// CFC twin of T_SafeTof_Tests: the same tests drawn as CFC diagrams, the way a TwinSAFE project is authored.
    FUNCTION_BLOCK T_SafeTof_Tests_CFC EXTENDS T_SafeCfcTestSuite
    VAR
    // Test_OutputDelayedOff
    group_1 : T_SafeGroup;
    fb_1 : T_SafeTof(group := group_1) := (Parameters := (DelayTime := T#100MS));
    trigStart_1 : R_TRIG;
    t0_1 : TON;
    t1_1 : TON;
    trig0_1 : R_TRIG;
    trig1_1 : R_TRIG;
END_VAR

Test_OutputDelayedOff();

METHOD PRIVATE Test_OutputDelayedOff
// note: this text did not pass the execution check against the stored diagram
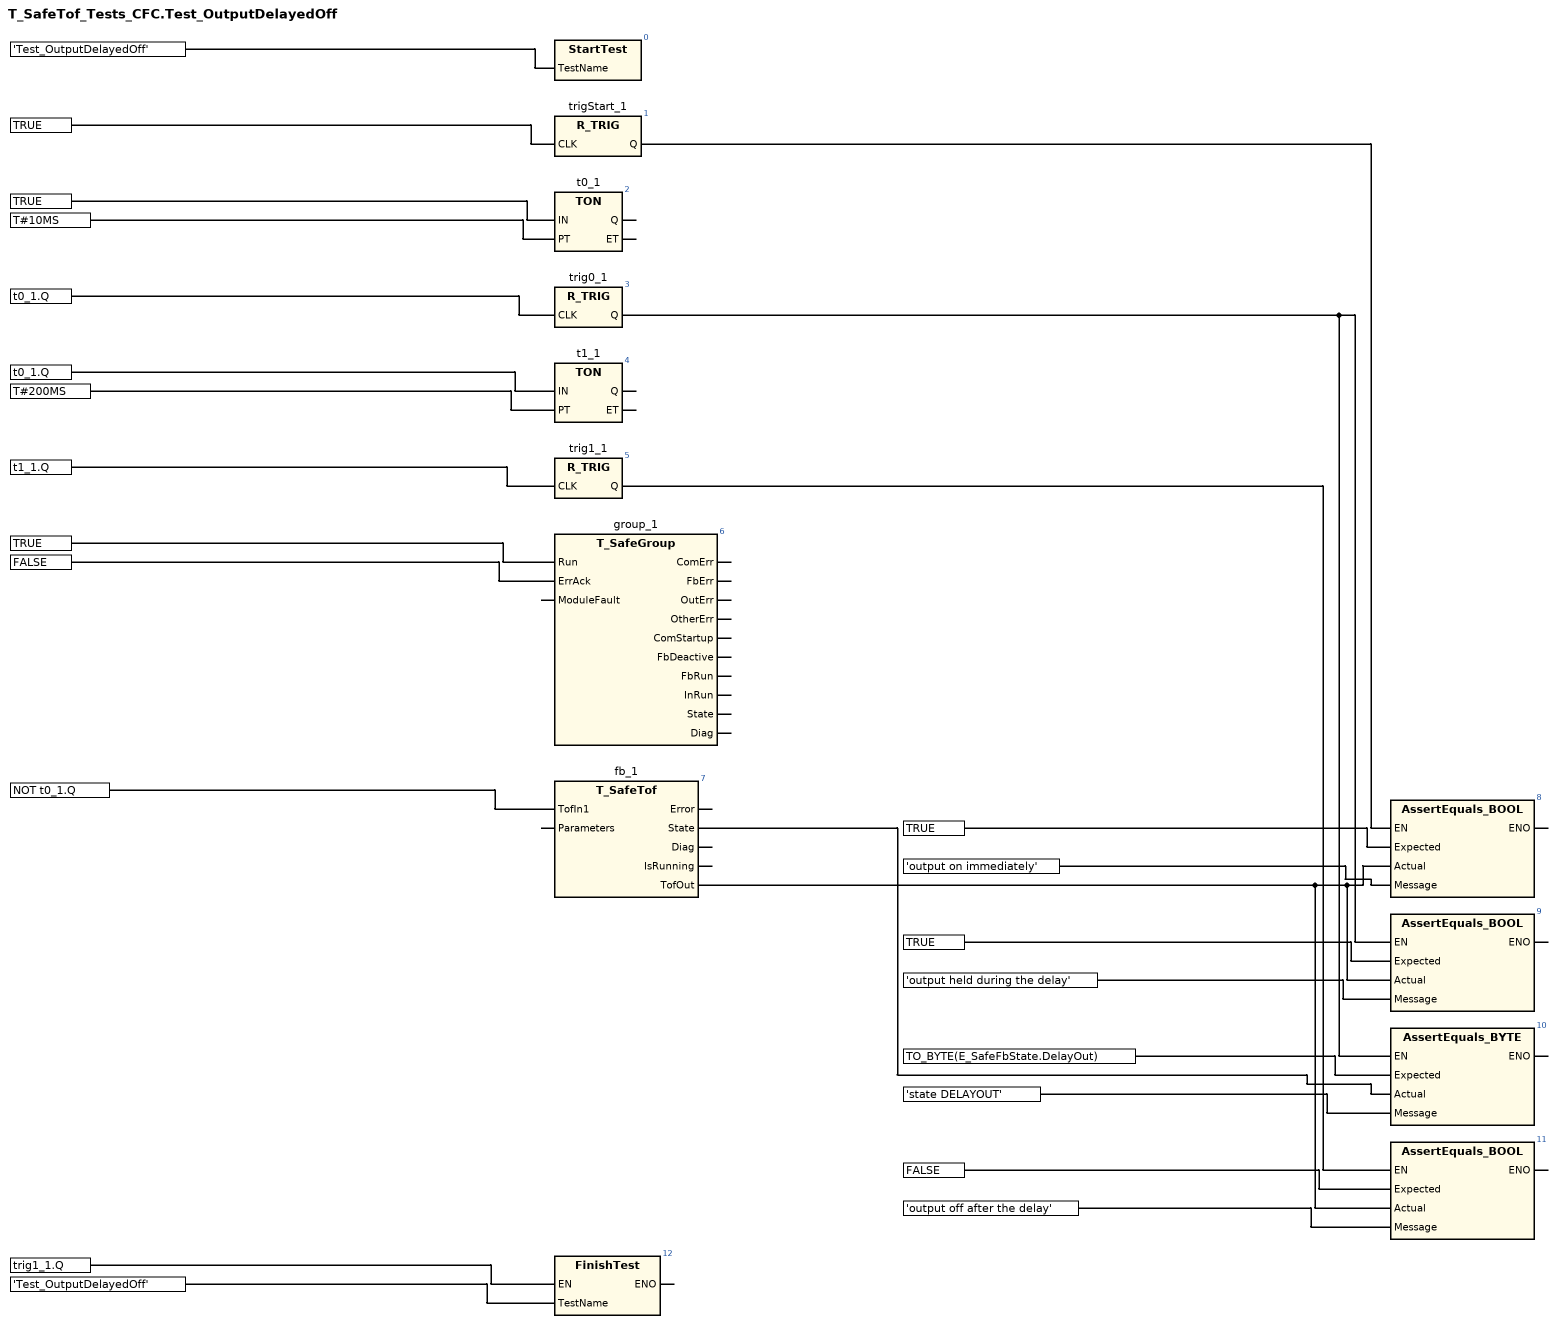
StartTest(TestName := 'Test_OutputDelayedOff');
trigStart_1(CLK := TRUE); // R_TRIG
t0_1(IN := TRUE, PT := T#10MS); // TON
trig0_1(CLK := t0_1.Q); // R_TRIG
t1_1(IN := t0_1.Q, PT := T#200MS); // TON
trig1_1(CLK := t1_1.Q); // R_TRIG
group_1(Run := TRUE, ErrAck := FALSE); // T_SafeGroup
fb_1(TofIn1 := NOT t0_1.Q); // T_SafeTof
IF trigStart_1.Q THEN AssertEquals_BOOL(Expected := TRUE, Actual := fb_1.TofOut, Message := 'output on immediately'); END_IF
IF trig0_1.Q THEN AssertEquals_BOOL(Expected := TRUE, Actual := fb_1.TofOut, Message := 'output held during the delay'); END_IF
IF trig0_1.Q THEN AssertEquals_BYTE(Expected := TO_BYTE(E_SafeFbState.DelayOut), Actual := fb_1.State, Message := 'state DELAYOUT'); END_IF
IF trig1_1.Q THEN AssertEquals_BOOL(Expected := FALSE, Actual := fb_1.TofOut, Message := 'output off after the delay'); END_IF
IF trig1_1.Q THEN FinishTest(TestName := 'Test_OutputDelayedOff'); END_IF
END_METHOD

END_FUNCTION_BLOCK

(* stored: Version 1.1.0.1, ProductVersion 3.1.4026.22
   POU T_SafeTof_Tests_CFC: Id {946bbad3-1e7e-527d-bd6b-28ed536bff55}, SpecialFunc None
   Method Test_OutputDelayedOff: Id {855a937f-e3c4-5a9e-85b3-cc9e76ea3486} *)
